DATA_BLOCK "StationData"
{ S7_Optimized_Access := 'TRUE' }
VERSION : 0.1
NON_RETAIN
"Station"

BEGIN

END_DATA_BLOCK

